Staubli VAL3: simulateHome.pgx

public program simulateHome()
  local bool l_bResult
  local bool l_bExit
begin
  if !rs:bIsCycle and workingMode()==1
    l_bResult=userPageConfirm("是否移动到Home位置？")
    if l_bResult
      rs:bSimulate=true

      taskCreate "simulate",50,goHome()
      sMsg="回Home过程。。。"
      call simulate_UI()
    endIf
  else
    userPageAlert("条件不满足：不再生产周期&切换到手动模式")
  endIf
end
